{attribute 'qualified_only'}
{attribute 'strict'}
{attribute 'to_string'}
TYPE E_PuckLockerState :
(
	Disabled                       := 0,
    WaitingForPuck                  := 10,
    LockingPuck                     := 20,
    Locked                          := 30,
    WaitingForPartRemoval           := 35,
    ReleasingPuck                   := 40,
    UnexpectedPuckRemovalFault      := 99
);
END_TYPE

(* stored: Version 1.1.0.1
   DUT E_PuckLockerState: Id {4b99b812-1afa-4a05-a159-d38479221f13} *)
